(* IEC 61131-3 sources: kns-port-domestic/tools/tests/fixtures/lowering/src/DUTs, 2 files *)

(* ---- ST_Cfg.dut.st ---- *)
// Настройки: массив структур с константой в границе
TYPE ST_Cfg :
STRUCT
    astSlot : ARRAY[0..GVL_Const.SLOTS_MAX - 1] OF ST_Slot;
END_STRUCT
END_TYPE

(* ---- ST_Slot.dut.st ---- *)
// Слот: массив в поле структуры с начальным значением, длина строки — константа
TYPE ST_Slot :
STRUCT
    xEnable : BOOL;
    rValue : REAL;
    arStep : ARRAY[1..4] OF REAL := [0.5, 1.0, 1.5, 2.0];
    sName : STRING(GVL_Const.NAME_LEN);
END_STRUCT
END_TYPE
